(* IEC 61131-3 sources: SortJet_MasterSPS_Aufbau.fbsproj/07_Auftragsverwaltung/Job_Stationen.prg.st^, 8 files *)

(* ---- Auftraege.act.st ---- *)
(* METADATA
{
	"v3Meta": {
		"objectGuid": "798febcb-6f60-456b-b36c-821ba17e31fa"
	}
}
*)
ACTION Auftraege
//-------------------------------------------------------------------------------------------------
// AUFTRAEGE: M_SB0_MMI_SortierungInputInQueue
//-------------------------------------------------------------------------------------------------
(* Hinweis:
   - Anlegetische \ Anlegewaende \ etc. mit einem Auftrag versehen
*)
IF ( M_SB0_MMI_SortierungInputInQueue ) THEN

  CASE tMmi2SpsInfo.wSortierungsInputInQueueStationNr OF

    cERSTE_STATION..cLETZTE_STATION:
      AuftragsSpeicherWand[tMmi2SpsInfo.wSortierungsInputInQueueStationNr, cWAND_1].NeuerAuftrag.rAuftragsHoehe       := tMmi2SpsInfo.rInputInQueueHoehe;
      AuftragsSpeicherWand[tMmi2SpsInfo.wSortierungsInputInQueueStationNr, cWAND_1].NeuerAuftrag.rAuftragsLaenge      := tMmi2SpsInfo.rInputInQueueLaenge;
      AuftragsSpeicherWand[tMmi2SpsInfo.wSortierungsInputInQueueStationNr, cWAND_1].NeuerAuftrag.rAuftragsDicke       := tMmi2SpsInfo.rInputInQueueDicke;
      AuftragsSpeicherWand[tMmi2SpsInfo.wSortierungsInputInQueueStationNr, cWAND_1].NeuerAuftrag.bLetzteScheibe       := 1;
      AuftragsSpeicherWand[tMmi2SpsInfo.wSortierungsInputInQueueStationNr, cWAND_1].NeuerAuftrag.wStationsNr          := tMmi2SpsInfo.wSortierungsInputInQueueStationNr;
      AuftragsSpeicherWand[tMmi2SpsInfo.wSortierungsInputInQueueStationNr, cWAND_1].NeuerAuftrag.wTransferwand        := tMmi2SpsInfo.wSlotZielStation;
      AuftragsSpeicherWand[tMmi2SpsInfo.wSortierungsInputInQueueStationNr, cWAND_1].NeuerAuftrag.wAnzahlScheiben      := 1; // es ist immer nur eine Scheibe anzulegen !
      AuftragsSpeicherWand[tMmi2SpsInfo.wSortierungsInputInQueueStationNr, cWAND_1].NeuerAuftrag.bErsteScheibe        := 1;
      AuftragsSpeicherWand[tMmi2SpsInfo.wSortierungsInputInQueueStationNr, cWAND_1].NeuerAuftrag.bModell              := tMmi2SpsInfo.wModellStatus.0;
      AuftragsSpeicherWand[tMmi2SpsInfo.wSortierungsInputInQueueStationNr, cWAND_1].NeuerAuftrag.rModellVersatzVorne  := tMmi2SpsInfo.rModellVersatzVorne;
      AuftragsSpeicherWand[tMmi2SpsInfo.wSortierungsInputInQueueStationNr, cWAND_1].NeuerAuftrag.rModellVersatzHinten := tMmi2SpsInfo.rModellversatzHinten;
      AuftragsSpeicherWand[tMmi2SpsInfo.wSortierungsInputInQueueStationNr, cWAND_1].NeuerAuftrag.wTransferstationsNr1 := tMmi2SpsInfo.wSourceTable;

      AuftragsSpeicherWand[tMmi2SpsInfo.wSortierungsInputInQueueStationNr, cWAND_1].NeuerAuftrag.wAuftrag := eStation_Anlegen;
      AuftragsSpeicherWand[tMmi2SpsInfo.wSortierungsInputInQueueStationNr, cWAND_1](bpNeuerAuftrag:=TRUE);

      M_SB0_MMI_SortierungInputInQueue := FALSE;

  END_CASE

END_IF

//-------------------------------------------------------------------------------------------------
// AUFTRAEGE: M_SB0_MMI_SORTIERUNGCANCELQUEUEDATA
//-------------------------------------------------------------------------------------------------
(* Hinweis:
   - Aktiven Auftrag eines Anlegetisches loeschen
*)
IF ( M_SB0_MMI_SORTIERUNGCANCELQUEUEDATA ) THEN

  (* Hinweis:
     - Dieser Auftrag darf nur im Automatik- Betrieb validiert \ bearbeitet werden
       => Sendet die HMI diesen Befehl z.B. im Handbetrieb würde der Merker fuer den Abbruch des Anlegeauftrags gesetzt und beim wechsel in den Automatikbetrieb
          würde der nächste Auftrag dann geloescht bzw. abgebrochen und damit verworfen.
       WICHTIG:
     - Sicherstellen das die Stationen diesem Automatikkreis auch angehoehren
  *)
  CASE tMmi2SpsInfo.wDeleteStationNr OF

    cERSTE_STATION..cLETZTE_STATION:
      IF NOT AutomatikAktiv(tMmi2SpsInfo.wDeleteStationNr) THEN
        M_SB0_MMI_SORTIERUNGCANCELQUEUEDATA := FALSE;
      ELSE

        IF ( AuftragsdatenWand[tMmi2SpsInfo.wDeleteStationNr, cWAND_1].wAuftrag = eStation_Anlegen ) THEN
          AuftragsdatenWand[tMmi2SpsInfo.wDeleteStationNr, cWAND_1].wAuftrag := eStation_Kein_Auftrag;
          Anlegen[tMmi2SpsInfo.wDeleteStationNr, cWAND_1](bpReset:=TRUE);
        ELSIF ( AuftragsdatenWand[tMmi2SpsInfo.wDeleteStationNr, cWAND_1].wAuftrag = eStation_Hoehenmessung ) THEN
          AuftragsdatenWand[tMmi2SpsInfo.wDeleteStationNr, cWAND_1].wAuftrag := eStation_Kein_Auftrag;
          Glashoehenmessung[tMmi2SpsInfo.wDeleteStationNr, cWAND_1](bpReset:=TRUE);
        ELSIF ( AuftragsdatenWand[tMmi2SpsInfo.wDeleteStationNr, cWAND_1].wAuftrag = eStation_Messfahrt ) THEN
          AuftragsdatenWand[tMmi2SpsInfo.wDeleteStationNr, cWAND_1].wAuftrag := eStation_Kein_Auftrag;
          Glaslaengenmessung[tMmi2SpsInfo.wDeleteStationNr, cWAND_1](bpReset:=TRUE);
        ELSE
          abpAbbruchAnlegeauftrag[tMmi2SpsInfo.wDeleteStationNr] := TRUE;
        END_IF

        M_SB0_MMI_SORTIERUNGCANCELQUEUEDATA := FALSE;

      END_IF

  END_CASE

END_IF

//-------------------------------------------------------------------------------------------------
// AUFTRAG: M_SB0_MMI_SHEET_ORDER_STATION
//-------------------------------------------------------------------------------------------------
(* Hinweis:
   - -
*)
IF ( M_SB0_MMI_SHEET_ORDER_STATION ) THEN

  IF ( tMmi2SpsInfo.wAuftragsWand = 0 ) THEN // WORKAROUND MMI
    tMmi2SpsInfo.wAuftragsWand := 1;
  END_IF
  IF ( tMmi2SpsInfo.wTransferwand = 0 ) THEN // WORKAROUND MMI
    tMmi2SpsInfo.wTransferwand := 1;
  END_IF

  CASE tMmi2SpsInfo.wStationsNr OF

    cERSTE_STATION..cLETZTE_STATION:
      AuftragsSpeicherWand[tMmi2SpsInfo.wStationsNr, tMmi2SpsInfo.wAuftragsWand].NeuerAuftrag.bModell                 := FALSE;

      AuftragsSpeicherWand[tMmi2SpsInfo.wStationsNr, tMmi2SpsInfo.wAuftragsWand].NeuerAuftrag.wStationsNr             := tMmi2SpsInfo.wStationsNr;          // Stationswand der Quellstation
      AuftragsSpeicherWand[tMmi2SpsInfo.wStationsNr, tMmi2SpsInfo.wAuftragsWand].NeuerAuftrag.wStationsWand           := tMmi2SpsInfo.wAuftragsWand;        // Stationswand der Quellstation
      AuftragsSpeicherWand[tMmi2SpsInfo.wStationsNr, tMmi2SpsInfo.wAuftragsWand].NeuerAuftrag.rStationsZielposition   := tMmi2SpsInfo.rStationsPosition;    // Stationsposition der Quellstation
      AuftragsSpeicherWand[tMmi2SpsInfo.wStationsNr, tMmi2SpsInfo.wAuftragsWand].NeuerAuftrag.rAuftragsLaenge         := tMmi2SpsInfo.rAuftragsLaenge;      // Länge der Scheibe/Batch
      AuftragsSpeicherWand[tMmi2SpsInfo.wStationsNr, tMmi2SpsInfo.wAuftragsWand].NeuerAuftrag.rAuftragsHoehe          := tMmi2SpsInfo.rAuftragsHoehe;       // Höhe der Scheibe/Batch
      AuftragsSpeicherWand[tMmi2SpsInfo.wStationsNr, tMmi2SpsInfo.wAuftragsWand].NeuerAuftrag.rAuftragsDicke          := tMmi2SpsInfo.rAuftragsDicke;       // Dicke der Scheibe/Batch
      AuftragsSpeicherWand[tMmi2SpsInfo.wStationsNr, tMmi2SpsInfo.wAuftragsWand].NeuerAuftrag.wErsteLetzteScheibe     := tMmi2SpsInfo.wErsteLetzteScheibe;  // Kennzeichnung Erste und Letzte Scheibe
      AuftragsSpeicherWand[tMmi2SpsInfo.wStationsNr, tMmi2SpsInfo.wAuftragsWand].NeuerAuftrag.wAnzahlScheiben         := tMmi2SpsInfo.wAnzahlScheiben;      // Anzahl der Scheiben
      AuftragsSpeicherWand[tMmi2SpsInfo.wStationsNr, tMmi2SpsInfo.wAuftragsWand].NeuerAuftrag.wTransferstationsNr1    := tMmi2SpsInfo.wTransferstationsNr1; // Stationsnummer der Zielstation 1
      AuftragsSpeicherWand[tMmi2SpsInfo.wStationsNr, tMmi2SpsInfo.wAuftragsWand].NeuerAuftrag.wTransferstationsNr2    := tMmi2SpsInfo.wTransferstationsNr2; // Stationsnummer der Zielstation 2
      AuftragsSpeicherWand[tMmi2SpsInfo.wStationsNr, tMmi2SpsInfo.wAuftragsWand].NeuerAuftrag.rTransferposition1      := tMmi2SpsInfo.rTransferposition1;   // Stationsposition der Zielstation 1
      AuftragsSpeicherWand[tMmi2SpsInfo.wStationsNr, tMmi2SpsInfo.wAuftragsWand].NeuerAuftrag.rTransferposition2      := tMmi2SpsInfo.rTransferposition2;   // Stationsposition der Zielstation 2
      AuftragsSpeicherWand[tMmi2SpsInfo.wStationsNr, tMmi2SpsInfo.wAuftragsWand].NeuerAuftrag.wTransferwand           := tMmi2SpsInfo.wTransferwand;        // Stationswand der Zielstationen
      AuftragsSpeicherWand[tMmi2SpsInfo.wStationsNr, tMmi2SpsInfo.wAuftragsWand].NeuerAuftrag.stAuftragsInformationen.wAuftragsInformationen  := tMmi2SpsInfo.wAuftragsTyp;         // Informationen zum Auftrag: Bit 1: Ein-Aus-Transport | Bit 2: Station entladen | Bit 3: Ziel FW | Bit 4-7: Wand entladen | etc.

      AuftragsSpeicherWand[tMmi2SpsInfo.wStationsNr, tMmi2SpsInfo.wAuftragsWand].NeuerAuftrag.rModellVersatzVorne     := tMmi2SpsInfo.rModellVersatzVorne;
      AuftragsSpeicherWand[tMmi2SpsInfo.wStationsNr, tMmi2SpsInfo.wAuftragsWand].NeuerAuftrag.rModellVersatzHinten    := tMmi2SpsInfo.rModellversatzHinten;

      IF ((tMmi2SpsInfo.rModellVersatzVorne > 0) OR (tMmi2SpsInfo.rModellVersatzHinten > 0 ) ) THEN
        AuftragsSpeicherWand[tMmi2SpsInfo.wStationsNr, tMmi2SpsInfo.wAuftragsWand].NeuerAuftrag.bModell              := TRUE;
      END_IF

      (* Hinweis:
         - Zuweisung der Bits "erste" und "letzte" Scheibe
      *)

      ErsteUndLetzteScheibeBits( wpErsteUndLetzteScheibe:= tMmi2SpsInfo.wErsteLetzteScheibe ,
                                 wpLetzteScheibe => wlLetzteScheibe,
                                 wpErsteScheibe  => wlErsteScheibe );

      AuftragsSpeicherWand[tMmi2SpsInfo.wStationsNr, tMmi2SpsInfo.wAuftragsWand].NeuerAuftrag.bLetzteScheibe  := wlLetzteScheibe > 0;  // Stationsposition der Zielstation 2
      AuftragsSpeicherWand[tMmi2SpsInfo.wStationsNr, tMmi2SpsInfo.wAuftragsWand].NeuerAuftrag.bErsteScheibe   := wlErsteScheibe  > 0;  // Stationswand der Zielstationen

      IF ( tMmi2SpsInfo.wAuftragsTyp.0 ) THEN
        AuftragsSpeicherWand[tMmi2SpsInfo.wStationsNr, tMmi2SpsInfo.wAuftragsWand].NeuerAuftrag.wAuftrag := eStation_Austransport;
      ELSE
        AuftragsSpeicherWand[tMmi2SpsInfo.wStationsNr, tMmi2SpsInfo.wAuftragsWand].NeuerAuftrag.wAuftrag := eStation_Eintransport;
      END_IF

      AuftragsSpeicherWand[tMmi2SpsInfo.wStationsNr, tMmi2SpsInfo.wAuftragsWand]( bpNeuerAuftrag := TRUE );

      M_SB0_MMI_SHEET_ORDER_STATION := FALSE;

    cERSTE_FREMDANLAGE_AUSLAUF..cLETZTE_FREMDANLAGE_EINLAUF:
      Job_Fremdanlage.AuftragsSpeicherFremdanlage[tMmi2SpsInfo.wStationsNr].NeuerAuftrag.wStationsNr            := tMmi2SpsInfo.wStationsNr;          // Stationswand der Quellstation
      Job_Fremdanlage.AuftragsSpeicherFremdanlage[tMmi2SpsInfo.wStationsNr].NeuerAuftrag.wStationsWand          := tMmi2SpsInfo.wAuftragsWand;        // Stationswand der Quellstation
      Job_Fremdanlage.AuftragsSpeicherFremdanlage[tMmi2SpsInfo.wStationsNr].NeuerAuftrag.rStationsZielposition  := tMmi2SpsInfo.rStationsPosition;    // Stationsposition der Quellstation
      Job_Fremdanlage.AuftragsSpeicherFremdanlage[tMmi2SpsInfo.wStationsNr].NeuerAuftrag.rAuftragsLaenge        := tMmi2SpsInfo.rAuftragsLaenge;      // Länge der Scheibe/Batch
      Job_Fremdanlage.AuftragsSpeicherFremdanlage[tMmi2SpsInfo.wStationsNr].NeuerAuftrag.rAuftragsHoehe         := tMmi2SpsInfo.rAuftragsHoehe;       // Höhe der Scheibe/Batch
      Job_Fremdanlage.AuftragsSpeicherFremdanlage[tMmi2SpsInfo.wStationsNr].NeuerAuftrag.rAuftragsDicke         := tMmi2SpsInfo.rAuftragsDicke;       // Dicke der Scheibe/Batch
      Job_Fremdanlage.AuftragsSpeicherFremdanlage[tMmi2SpsInfo.wStationsNr].NeuerAuftrag.wErsteLetzteScheibe    := tMmi2SpsInfo.wErsteLetzteScheibe;  // Kennzeichnung Erste und Letzte Scheibe
      Job_Fremdanlage.AuftragsSpeicherFremdanlage[tMmi2SpsInfo.wStationsNr].NeuerAuftrag.wAnzahlScheiben        := tMmi2SpsInfo.wAnzahlScheiben;      // Anzahl der Scheiben
      Job_Fremdanlage.AuftragsSpeicherFremdanlage[tMmi2SpsInfo.wStationsNr].NeuerAuftrag.wTransferstationsNr1   := tMmi2SpsInfo.wTransferstationsNr1; // Stationsnummer der Zielstation 1
      Job_Fremdanlage.AuftragsSpeicherFremdanlage[tMmi2SpsInfo.wStationsNr].NeuerAuftrag.wTransferstationsNr2   := tMmi2SpsInfo.wTransferstationsNr2; // Stationsnummer der Zielstation 2
      Job_Fremdanlage.AuftragsSpeicherFremdanlage[tMmi2SpsInfo.wStationsNr].NeuerAuftrag.rTransferposition1     := tMmi2SpsInfo.rTransferposition1;   // Stationsposition der Zielstation 1
      Job_Fremdanlage.AuftragsSpeicherFremdanlage[tMmi2SpsInfo.wStationsNr].NeuerAuftrag.rTransferposition2     := tMmi2SpsInfo.rTransferposition2;   // Stationsposition der Zielstation 2
      Job_Fremdanlage.AuftragsSpeicherFremdanlage[tMmi2SpsInfo.wStationsNr].NeuerAuftrag.wTransferwand          := tMmi2SpsInfo.wTransferwand;        // Stationswand der Zielstationen
      Job_Fremdanlage.AuftragsSpeicherFremdanlage[tMmi2SpsInfo.wStationsNr].NeuerAuftrag.stAuftragsInformationen.wAuftragsInformationen := tMmi2SpsInfo.wAuftragsTyp;         // Informationen zum Auftrag: Bit 1: Ein-Aus-Transport | Bit 2: Station entladen | Bit 3: Ziel FW | Bit 4-7: Wand entladen | etc.

      Job_Fremdanlage.AuftragsSpeicherFremdanlage[tMmi2SpsInfo.wStationsNr].NeuerAuftrag.rModellVersatzVorne  := tMmi2SpsInfo.rModellVersatzVorne;
      Job_Fremdanlage.AuftragsSpeicherFremdanlage[tMmi2SpsInfo.wStationsNr].NeuerAuftrag.rModellVersatzHinten := tMmi2SpsInfo.rModellversatzHinten;

      IF ((tMmi2SpsInfo.rModellVersatzVorne > 0) OR (tMmi2SpsInfo.rModellVersatzHinten > 0 ) ) THEN
        Job_Fremdanlage.AuftragsSpeicherFremdanlage[tMmi2SpsInfo.wStationsNr].NeuerAuftrag.bModell              := TRUE;
      END_IF

      (* Hinweis:
         - Zuweisung der Bits "erste" und "letzte" Scheibe
      *)
      ErsteUndLetzteScheibeBits( wpErsteUndLetzteScheibe:= tMmi2SpsInfo.wErsteLetzteScheibe ,
                                 wpLetzteScheibe => wlLetzteScheibe,
                                 wpErsteScheibe  => wlErsteScheibe );

      Job_Fremdanlage.AuftragsSpeicherFremdanlage[tMmi2SpsInfo.wStationsNr].NeuerAuftrag.bLetzteScheibe  := wlLetzteScheibe > 0;  // Stationsposition der Zielstation 2
      Job_Fremdanlage.AuftragsSpeicherFremdanlage[tMmi2SpsInfo.wStationsNr].NeuerAuftrag.bErsteScheibe   := wlErsteScheibe  > 0;  // Stationswand der Zielstationen

      IF ( tMmi2SpsInfo.wAuftragsTyp.0 ) THEN
        Job_Fremdanlage.AuftragsSpeicherFremdanlage[tMmi2SpsInfo.wStationsNr].NeuerAuftrag.wAuftrag := eStation_Austransport;
      ELSE
        Job_Fremdanlage.AuftragsSpeicherFremdanlage[tMmi2SpsInfo.wStationsNr].NeuerAuftrag.wAuftrag := eStation_Eintransport;
      END_IF

      Job_Fremdanlage.AuftragsSpeicherFremdanlage[tMmi2SpsInfo.wStationsNr]( bpNeuerAuftrag := TRUE );

      M_SB0_MMI_SHEET_ORDER_STATION := FALSE;

    ELSE

      M_SB0_MMI_SHEET_ORDER_STATION := FALSE;

      wpgFehlerdaten[0] := tMmi2SpsInfo.wStationsNr;
      wpgFehlerdaten[1] := tMmi2SpsInfo.wAuftragsWand;
      SpsError( eFehler_Station,
                cMELDUNG_AUFTRAGSDATEN_UNGUELTIGE_STATION,
                tMmi2SpsInfo.wStationsNr,
                AutomatikkreisBestimmen(tMmi2SpsInfo.wStationsNr),
                wpgFehlerdaten );

  END_CASE

END_IF

//-------------------------------------------------------------------------------------------------
// AUFTRAG: M_SB0_MMI_MEASSURERESULT
//-------------------------------------------------------------------------------------------------
(* Hinweis:
   - Scheibeneinlauffreigabe für Anlegetisch
     => Gilt fuer Stationen mit einem Scanner
*)
IF ( M_SB0_MMI_MEASSURERESULT ) THEN

  M_SB0_MMI_MEASSURERESULT := FALSE;

  CASE (tMmi2SpsInfo.wMmiNummerAnlegeStation) OF

    cERSTE_STATION..cLETZTE_STATION:
      ;
    //Anlegewand202.bpFreigabeScheibe      := (tMmi2SpsInfo.wFreigabe = 1);
    //Anlegewand202.bpKeineFreigabeScheibe := (tMmi2SpsInfo.wFreigabe = 0);

    ELSE
      wpgFehlerdaten[0]:= tMmi2SpsInfo.wMmiNummerAnlegeStation;
      wpgFehlerdaten[1]:= tMmi2SpsInfo.wFreigabeStation;
      SpsError( eFehler_Station,
                cMELDUNG_SCANNER_NACHRICHT_FALSCHE_STATION,
                tMmi2SpsInfo.wMmiNummerAnlegeStation,
                AutomatikkreisBestimmen(tMmi2SpsInfo.wMmiNummerAnlegeStation),
                wpgFehlerdaten );

  END_CASE

END_IF

//-------------------------------------------------------------------------------------------------
// AUFTRAG: M_SB0_MMI_STATIONSTATUS
//-------------------------------------------------------------------------------------------------
IF ( M_SB0_MMI_STATIONSTATUS ) THEN

  M_SB0_MMI_STATIONSTATUS := FALSE;

  CASE tMmi2SpsInfo.wStationsNummer OF

    // -------------------------------------------------------------------
    cERSTE_STATION..cLETZTE_STATION:
      (* Hinweis:
         - Aktivieren / Deaktivieren der Station
      *)
      starrStationBasisParameter[tMmi2SpsInfo.wStationsNummer].stMKs.bDeaktivieren := ( NOT tMmi2SpsInfo.wStationsStatusWord7.0 );

    // -------------------------------------------------------------------
    cERSTES_SHUTTLE..cLETZTES_SHUTTLE:
      (* Hinweis:
         - Aktivieren / Deaktivieren der Station
      *)
      starrShuttleBasisParameter[tMmi2SpsInfo.wStationsNummer].stMKs.bDeaktivieren := ( NOT tMmi2SpsInfo.wStationsStatusWord7.0 );

    // -------------------------------------------------------------------
    cERSTES_TRANSFERSHUTTLE..cLETZTES_TRANSFERSHUTTLE:
      (* Hinweis:
         - Aktivieren / Deaktivieren der Station
      *)
      starrTransfershuttleBasisParameter[tMmi2SpsInfo.wStationsNummer].stMKs.bDeaktivieren := ( NOT tMmi2SpsInfo.wStationsStatusWord7.0 );

    // -------------------------------------------------------------------
    cERSTE_FAECHERWAGENSTATIONS_NR..cLETZTE_FAECHERWAGENSTATIONS_NR:
      (* Hinweis:
         - Aktivieren / Deaktivieren der Station
      *)
      starrFaecherwagenBasisParameter[tMmi2SpsInfo.wStationsNummer].stMKs.bDeaktivieren := ( NOT tMmi2SpsInfo.wStationsStatusWord7.0 );
      aFaecherwagenstation[tMmi2SpsInfo.wStationsNummer].wRFID_Nummer_Schreiben := tMmi2SpsInfo.wStationsStatusWord8;

      // Statuswort 1 Bit 0: bei Faecherwagenstationen loest es den Sicherheitskreis-Reset der Station aus
      // (Sicherheitsrelais der Station quittieren)
      IF ( tMmi2SpsInfo.wStationsStatusWord1.0 ) THEN
        aFaecherwagenstation[tMmi2SpsInfo.wStationsNummer].bStarteSicherheitskreisReset := TRUE;
      END_IF

    // -------------------------------------------------------------------
    ELSE
      wpgFehlerdaten[0] := tMmi2SpsInfo.wStationsNummer;
      wpgFehlerdaten[1] := tMmi2SpsInfo.wStationsStatusWord5;
      SpsHinweis( eFehler_Mmi,
                  cMELDUNG_MMI_AUFTRAGSDATEN_UNGUELTIGE_STATIONSNUMMER,
                  0,
                  AutomatikkreisBestimmen(0),
                  wpgFehlerdaten );

  END_CASE

END_IF

//-------------------------------------------------------------------------------------------------
// AUFTRAG: M_SB0_MMI_REQUESTTILTSTATION
//-------------------------------------------------------------------------------------------------

(* Hinweis:
   - Auftrag zum leeren einer Station (Starten eines Austransports)
*)
IF ( M_SB0_MMI_REQUESTTILTSTATION ) THEN

  CASE tMmi2SpsInfo.wSortierungsInputSwingStationNr OF

    cERSTE_STATION..cLETZTE_STATION:
      AuftragsSpeicherWand[tMmi2SpsInfo.wSortierungsInputSwingStationNr, cWAND_1].NeuerAuftrag.wAuftrag      := eStation_Vortransport;
      AuftragsSpeicherWand[tMmi2SpsInfo.wSortierungsInputSwingStationNr, cWAND_1].NeuerAuftrag.wStationsNr   := tMmi2SpsInfo.wSortierungsInputSwingStationNr;
      AuftragsSpeicherWand[tMmi2SpsInfo.wSortierungsInputSwingStationNr, cWAND_1].NeuerAuftrag.wStationsWand := cWAND_1;
      AuftragsSpeicherWand[tMmi2SpsInfo.wSortierungsInputSwingStationNr, cWAND_1]( bpNeuerAuftrag := TRUE );

    ELSE
      wpgFehlerdaten[0] := tMmi2SpsInfo.wSortierungsInputSwingStationNr;
      SpsHinweis( eFehler_Mmi,
                  cMELDUNG_MMI_AUFTRAGSDATEN_UNGUELTIGE_STATIONSNUMMER,
                  0,
                  AutomatikkreisBestimmen(0),
                  wpgFehlerdaten );

  END_CASE

  M_SB0_MMI_REQUESTTILTSTATION := FALSE;

END_IF
END_ACTION

(* ---- Auftragsverwaltung.act.st ---- *)
(* METADATA
{
	"v3Meta": {
		"objectGuid": "ab37f234-5c30-423e-82fd-562034963c76"
	}
}
*)
ACTION Auftragsverwaltung
//-------------------------------------------------------------------------------------------------
// BAUSTEIN: AUFTRAGSVERWALTUNG
//-------------------------------------------------------------------------------------------------
FOR wlIndex := cERSTE_STATION TO cLETZTE_STATION DO

  AuftragsSpeicherStation[wlIndex]();

  IF AuftragsSpeicherStation[wlIndex].bpAuftragverfuegbar
     AND ( AuftragsdatenStation[wlIndex].wAuftrag = eStation_Kein_Auftrag
           OR AuftragsdatenStation[wlIndex].wAuftrag = eStation_Belegt
           OR AuftragsdatenStation[wlIndex].wAuftrag = eStation_Warte_Auf_Eintransport )
  THEN
    AuftragsSpeicherStation[wlIndex].bpNaechsterAuftrag := TRUE;
    AuftragsSpeicherStation[wlIndex]();
    AuftragsdatenStation[wlIndex] := AuftragsSpeicherStation[wlIndex].AktAuftrag;
  END_IF

  FOR wlIndexWand := cWAND_1 TO cANZAHL_WAENDE DO

    AuftragsSpeicherWand[wlIndex, wlIndexWand]();

    IF AuftragsSpeicherWand[wlIndex, wlIndexWand].bpAuftragverfuegbar
       AND ( AuftragsdatenWand[wlIndex, wlIndexWand].wAuftrag = eStation_Kein_Auftrag
             OR AuftragsdatenWand[wlIndex, wlIndexWand].wAuftrag = eStation_Belegt
             OR AuftragsdatenWand[wlIndex, wlIndexWand].wAuftrag = eStation_Warte_Auf_Eintransport
             OR AuftragsdatenWand[wlIndex, wlIndexWand].wAuftrag = eStation_Warte_Auf_Austransport  )
    THEN
      AuftragsSpeicherWand[wlIndex, wlIndexWand].bpNaechsterAuftrag := TRUE;
      AuftragsSpeicherWand[wlIndex, wlIndexWand]();
      AuftragsdatenWand[wlIndex, wlIndexWand] := AuftragsSpeicherWand[wlIndex, wlIndexWand].AktAuftrag;
    END_IF

  END_FOR

END_FOR
END_ACTION

(* ---- Reset.act.st ---- *)
(* METADATA
{
	"v3Meta": {
		"objectGuid": "37f6c3a9-3bba-4d57-9c53-2ef1e7be2c3a"
	}
}
*)
ACTION Reset
//-------------------------------------------------------------------------------------------------
// AKTION: RESET
//-------------------------------------------------------------------------------------------------

FOR wlIndexReset := cERSTER_AUTOMATIKKREIS TO cLETZTER_AUTOMATIKKREIS DO

  IF ( abpReset[wlIndexReset] ) THEN

    abpReset[wlIndexReset] := FALSE;
    abpFehler[wlIndexReset] := FALSE;

    FOR wlIndex := cERSTE_STATION TO cLETZTE_STATION DO

      IF StationInAutomatikkreis(starrStationBasisParameter[wlIndex].stMKs.eaAutomatikkreis, wlIndexReset) THEN

        abpAbbruchAnlegeauftrag[wlIndex] := FALSE;

        AuftragsSpeicherStation[wlIndex].bpReset := TRUE;
        AuftragsSpeicherStation[wlIndex]();

        AuftragsdatenStation[wlIndex].wAuftrag := eStation_Kein_Auftrag;

        starrStationBasisParameter[wlIndex].bReset := TRUE;

        FOR wlIndexWand := cWAND_1 TO cANZAHL_WAENDE DO

          AuftragsSpeicherWand[wlIndex,wlIndexWand].bpReset := TRUE;
          AuftragsSpeicherWand[wlIndex,wlIndexWand]();

          AuftragsdatenWand[wlIndex, wlIndexWand].wAuftrag := eStation_Kein_Auftrag;

          ailScheibenZuQuittierenEintransport[wlIndex, wlIndexWand] := 0;
          ailScheibenZuQuittierenAustransport[wlIndex, wlIndexWand] := 0;

          ablMerkerLetzteScheibeStation[wlIndex, wlIndexWand] := FALSE;

          ablFreigabeZurParalleleBausteinAnsteuerung[wlIndex,wlIndexWand] := FALSE;
          abpStarteParalleleBausteinAnsteuerung[wlIndex, wlIndexWand]     := FALSE;

        END_FOR

      END_IF

    END_FOR

  END_IF

END_FOR
END_ACTION

(* ---- Schnittstelle_Stationen.act.st ---- *)
(* METADATA
{
	"v3Meta": {
		"objectGuid": "2f0e1e2b-c489-43f6-919f-1d41b03fa1f2"
	}
}
*)
ACTION Schnittstelle_Stationen
//-------------------------------------------------------------------------------------------------
// SCHNITTSTELLE ZWISCHEN DEN STATIONEN
//-------------------------------------------------------------------------------------------------

//  KOPPLUNGEN

//starrFremdanlageEinlaufStationBasisParameter[501].InGlasTransportNachfolger[cWAND_1] := starrStationBasisParameter[cSTATION_201].OutGlasTransport[cWAND_1];
//starrStationBasisParameter[cSTATION_201].InGlasTransportVorgaenger[cWAND_1] := starrFremdanlageEinlaufStationBasisParameter[501].OutGlasTransport[cWAND_1];

FOR wlIndex := cERSTE_STATION TO cLETZTE_FREMDANLAGE_EINLAUF DO

  // Struktur für die Zielstation der Kopplung finden
  stLokaleKopplungZielStation REF= getBasis(wlIndex);

  IF __ISVALIDREF(stLokaleKopplungZielStation) THEN

    // Kopplung Vorgänger
    stLokaleKopplungsStation REF= getBasis(stLokaleKopplungZielStation.stMKs.stSchnittstellendaten.wVorgaengerStation);

    IF __ISVALIDREF(stLokaleKopplungsStation) THEN
      FOR wlIndexWand := cWAND_1 TO cANZAHL_WAENDE DO
        stLokaleKopplungZielStation.InGlasTransportVorgaenger[wlIndexWand] := stLokaleKopplungsStation.OutGlasTransport[cWAND_1];
      END_FOR
    END_IF

    // Kopplung Nachfolger
    stLokaleKopplungsStation REF= getBasis(stLokaleKopplungZielStation.stMKs.stSchnittstellendaten.wNachfolgerStation);

    IF __ISVALIDREF(stLokaleKopplungsStation) THEN
      FOR wlIndexWand := cWAND_1 TO cANZAHL_WAENDE DO
        stLokaleKopplungZielStation.InGlasTransportNachfolger[wlIndexWand] := stLokaleKopplungsStation.OutGlasTransport[cWAND_1];
      END_FOR
    END_IF

  END_IF

END_FOR
END_ACTION

(* ---- Station.meth.st ---- *)
(* METADATA
{
	"v3Meta": {
		"objectGuid": "6e43b8d4-0bae-4a3f-b309-8e06ab9993e4"
	}
}
*)
METHOD INTERNAL Station
VAR_INPUT
  wStation : WORD;
  wWand    : WORD;
END_VAR

// ****************************************************9*********************************************
// STEUERUNG: ANLEGEN
// *************************************************************************************************

IF ( AuftragsdatenWand[wStation, wWand].wAuftrag = eStation_Anlegen ) THEN
  (* Hinweis:
     - Aufruf der Schrittkette
  *)
  Anlegen[wStation, wWand]( Auftragsdaten := AuftragsdatenWand[wStation, wWand], bpAbbruchAnlegeauftrag := abpAbbruchAnlegeauftrag[wStation], wStation := wStation);
  (* Hinweis:
     - Abschluss der Schrittkette
  *)
  IF Anlegen[wStation, wWand].bpDone THEN
    abpAbbruchAnlegeauftrag[wStation] := FALSE;
    AuftragsdatenWand[wStation, wWand] := Anlegen[wStation, wWand].Auftragsdaten;
    Anlegen[wStation, wWand](bpReset := TRUE);
  END_IF
  (* Hinweis:
     - Fehler-Auswertung
  *)
  ablFehler[wStation, wWand] := Anlegen[wStation, wWand].bpFehler;
  IF rtlFehler[wStation, wWand].Q THEN
    AutomatikFehlerSetzen(starrStationBasisParameter[wStation].stMKs.eaAutomatikkreis, abpFehler);
  END_IF
ELSE
  (* Hinweis:
     - Reset der Schrittkette
  *)
  IF ( Anlegen[wStation, wWand].steplSchritt > STEP_0_E ) THEN
    Anlegen[wStation, wWand](bpReset := TRUE);
  END_IF
END_IF

// ****************************************************9*********************************************
// STEUERUNG: ABNEHMEN
// *************************************************************************************************

IF ( AuftragsdatenWand[wStation, wWand].wAuftrag = eStation_Abnehmen ) THEN
  (* Hinweis:
     - Aufruf der Schrittkette
  *)
  Abnehmen[wStation, wWand]( Auftragsdaten := AuftragsdatenWand[wStation, wWand], wStation := wStation);
  (* Hinweis:
     - Abschluss der Schrittkette
  *)
  IF Abnehmen[wStation, wWand].bpDone THEN
    abpAbbruchAnlegeauftrag[wStation] := FALSE;
    AuftragsdatenWand[wStation, wWand] := Abnehmen[wStation, wWand].Auftragsdaten;
    Abnehmen[wStation, wWand](bpReset := TRUE);
  END_IF
  (* Hinweis:
     - Fehler-Auswertung
  *)
  ablFehler[wStation, wWand] := Abnehmen[wStation, wWand].bpFehler;
  IF rtlFehler[wStation, wWand].Q THEN
    AutomatikFehlerSetzen(starrStationBasisParameter[wStation].stMKs.eaAutomatikkreis, abpFehler);
  END_IF
ELSE
  (* Hinweis:
     - Reset der Schrittkette
  *)
  IF ( Abnehmen[wStation, wWand].steplSchritt > STEP_0_E ) THEN
    Abnehmen[wStation, wWand](bpReset := TRUE);
  END_IF
END_IF

// ****************************************************9*********************************************
// STEUERUNG: HÖHENMESSUNG
// *************************************************************************************************

IF ( AuftragsdatenWand[wStation, wWand].wAuftrag = eStation_Hoehenmessung ) THEN
  (* Hinweis:
     - Aufruf der Schrittkette
  *)
  Glashoehenmessung[wStation, wWand]( Auftragsdaten := AuftragsdatenWand[wStation, wWand], wStation := wStation, bpAbbruchAnlegeauftrag := abpAbbruchAnlegeauftrag[wStation]);
  (* Hinweis:
     - Abschluss der Schrittkette
  *)
  IF Glashoehenmessung[wStation, wWand].bpDone THEN
    abpAbbruchAnlegeauftrag[wStation] := FALSE;
    AuftragsdatenWand[wStation, wWand] := Glashoehenmessung[wStation, wWand].Auftragsdaten;
    Glashoehenmessung[wStation, wWand](bpReset := TRUE);
  END_IF
  (* Hinweis:
     - Fehler-Auswertung
  *)
  ablFehler[wStation, wWand] := Glashoehenmessung[wStation, wWand].bpFehler;
  IF rtlFehler[wStation, wWand].Q THEN
    AutomatikFehlerSetzen(starrStationBasisParameter[wStation].stMKs.eaAutomatikkreis, abpFehler);
  END_IF
ELSE
  (* Hinweis:
     - Reset der Schrittkette
  *)
  IF ( Glashoehenmessung[wStation, wWand].steplSchritt > STEP_0_E ) THEN
    Glashoehenmessung[wStation, wWand](bpReset := TRUE);
  END_IF
END_IF

// ****************************************************9*********************************************
// STEUERUNG: LÄNGENMESSUNG
// *************************************************************************************************

IF ( AuftragsdatenWand[wStation, wWand].wAuftrag = eStation_Messfahrt ) THEN
  (* Hinweis:
     - Aufruf der Schrittkette
  *)
  Glaslaengenmessung[wStation, wWand]( Auftragsdaten := AuftragsdatenWand[wStation, wWand], wStation := wStation, bpAbbruchAnlegeauftrag := abpAbbruchAnlegeauftrag[wStation] );
  (* Hinweis:
     - Abschluss der Schrittkette
  *)
  IF Glaslaengenmessung[wStation, wWand].bpDone THEN
    abpAbbruchAnlegeauftrag[wStation] := FALSE;
    AuftragsdatenWand[wStation, wWand] := Glaslaengenmessung[wStation, wWand].Auftragsdaten;
    Glaslaengenmessung[wStation, wWand](bpReset := TRUE);
  END_IF
  (* Hinweis:
     - Fehler-Auswertung
  *)
  ablFehler[wStation, wWand] := Glaslaengenmessung[wStation, wWand].bpFehler;
  IF rtlFehler[wStation, wWand].Q THEN
    AutomatikFehlerSetzen(starrStationBasisParameter[wStation].stMKs.eaAutomatikkreis, abpFehler);
  END_IF
ELSE
  (* Hinweis:
     - Reset der Schrittkette
  *)
  IF ( Glaslaengenmessung[wStation, wWand].steplSchritt > STEP_0_E ) THEN
    Glaslaengenmessung[wStation, wWand](bpReset := TRUE);
  END_IF
END_IF

// ****************************************************9*********************************************
// STEUERUNG: Eintransport
// *************************************************************************************************

IF ( AuftragsdatenWand[wStation, wWand].wAuftrag = eStation_Eintransport ) THEN
  (* Hinweis:
     - Aufruf der Schrittkette
  *)
  Eintransport[wStation, wWand]( Auftragsdaten := AuftragsdatenWand[wStation, wWand], wStation := wStation, wWand := wWand);
  (* Hinweis:
     - Abschluss der Schrittkette
  *)
  IF Eintransport[wStation, wWand].bpDone THEN
    AuftragsdatenWand[wStation, wWand] := Eintransport[wStation, wWand].Auftragsdaten;
    Eintransport[wStation, wWand](bpReset := TRUE);
  END_IF
  (* Hinweis:
     - Fehler-Auswertung
  *)
  ablFehler[wStation, wWand] := Eintransport[wStation, wWand].bpFehler;
  IF rtlFehler[wStation, wWand].Q THEN
    AutomatikFehlerSetzen(starrStationBasisParameter[wStation].stMKs.eaAutomatikkreis, abpFehler);
  END_IF
ELSE
  (* Hinweis:
     - Reset der Schrittkette
  *)
  IF ( Eintransport[wStation, wWand].steplSchritt > STEP_0_E ) THEN
    Eintransport[wStation, wWand](bpReset := TRUE);
  END_IF
END_IF

// ****************************************************9*********************************************
// STEUERUNG: AUSTRANSPORT
// *************************************************************************************************

IF ( AuftragsdatenWand[wStation, wWand].wAuftrag = eStation_Austransport ) THEN
  (* Hinweis:
     - Aufruf der Schrittkette
  *)
  Austransport[wStation, wWand]( Auftragsdaten := AuftragsdatenWand[wStation, wWand], wStation := wStation, wWand := wWand);
  (* Hinweis:
     - Abschluss der Schrittkette
  *)
  IF Austransport[wStation, wWand].bpDone THEN
    AuftragsdatenWand[wStation, wWand] := Austransport[wStation, wWand].Auftragsdaten;
    Austransport[wStation, wWand](bpReset := TRUE);
  END_IF
  (* Hinweis:
     - Fehler-Auswertung
  *)
  ablFehler[wStation, wWand] := Austransport[wStation, wWand].bpFehler;
  IF rtlFehler[wStation, wWand].Q THEN
    AutomatikFehlerSetzen(starrStationBasisParameter[wStation].stMKs.eaAutomatikkreis, abpFehler);
  END_IF
ELSE
  (* Hinweis:
     - Reset der Schrittkette
  *)
  IF ( Austransport[wStation, wWand].steplSchritt > STEP_0_E ) THEN
    Austransport[wStation, wWand](bpReset := TRUE);
  END_IF
END_IF

// ****************************************************9*********************************************
// STEUERUNG: DURCHTRANSPORT
// *************************************************************************************************

IF ( AuftragsdatenWand[wStation, wWand].wAuftrag = eStation_Durchtransport ) THEN
  (* Hinweis:
     - Aufruf der Schrittkette
  *)
  Durchtransport[wStation, wWand]( Auftragsdaten := AuftragsdatenWand[wStation, wWand], wStation := wStation, wWand := wWand);
  (* Hinweis:
     - Abschluss der Schrittkette
  *)
  IF Durchtransport[wStation, wWand].bpDone THEN
    AuftragsdatenWand[wStation, wWand] := Durchtransport[wStation, wWand].Auftragsdaten;
    Durchtransport[wStation, wWand](bpReset := TRUE);
  END_IF
  (* Hinweis:
     - Fehler-Auswertung
  *)
  ablFehler[wStation, wWand] := Durchtransport[wStation, wWand].bpFehler;
  IF rtlFehler[wStation, wWand].Q THEN
    AutomatikFehlerSetzen(starrStationBasisParameter[wStation].stMKs.eaAutomatikkreis, abpFehler);
  END_IF
ELSE
  (* Hinweis:
     - Reset der Schrittkette
  *)
  IF ( Durchtransport[wStation, wWand].steplSchritt > STEP_0_E ) THEN
    Durchtransport[wStation, wWand](bpReset := TRUE);
  END_IF
END_IF

// ****************************************************9*********************************************
// STEUERUNG: Vortransport
// *************************************************************************************************

IF ( AuftragsdatenWand[wStation, wWand].wAuftrag = eStation_Vortransport ) THEN
  (* Hinweis:
     - Aufruf der Schrittkette
  *)
  Vortransport[wStation, wWand]( Auftragsdaten := AuftragsdatenWand[wStation, wWand], wStation := wStation, wWand := wWand);
  (* Hinweis:
     - Abschluss der Schrittkette
  *)
  IF Vortransport[wStation, wWand].bpDone THEN
    AuftragsdatenWand[wStation, wWand] := Vortransport[wStation, wWand].Auftragsdaten;
    Vortransport[wStation, wWand](bpReset := TRUE);
  END_IF
  (* Hinweis:
     - Fehler-Auswertung
  *)
  ablFehler[wStation, wWand] := Vortransport[wStation, wWand].bpFehler;
  IF rtlFehler[wStation, wWand].Q THEN
    AutomatikFehlerSetzen(starrStationBasisParameter[wStation].stMKs.eaAutomatikkreis, abpFehler);
  END_IF
ELSE
  (* Hinweis:
     - Reset der Schrittkette
  *)
  IF ( Vortransport[wStation, wWand].steplSchritt > STEP_0_E ) THEN
    Vortransport[wStation, wWand](bpReset := TRUE);
  END_IF
END_IF

// ****************************************************9*********************************************
// STEUERUNG: TRANSPORTKOPPLUNG
// *************************************************************************************************

IF ( AuftragsdatenWand[wStation, wWand].wAuftrag = eStation_Transportkopplung ) THEN
  (* Hinweis:
     - Aufruf der Schrittkette
  *)
  Transportkopplung[wStation, wWand]( Auftragsdaten := AuftragsdatenWand[wStation, wWand], wStation := wStation, wWand := wWand);
  (* Hinweis:
     - Abschluss der Schrittkette
  *)
  IF Transportkopplung[wStation, wWand].bpDone THEN
    AuftragsdatenWand[wStation, wWand] := Transportkopplung[wStation, wWand].Auftragsdaten;
    Transportkopplung[wStation, wWand](bpReset := TRUE);
  END_IF
  (* Hinweis:
     - Fehler-Auswertung
  *)
  ablFehler[wStation, wWand] := Transportkopplung[wStation, wWand].bpFehler;
  IF rtlFehler[wStation, wWand].Q THEN
    AutomatikFehlerSetzen(starrStationBasisParameter[wStation].stMKs.eaAutomatikkreis, abpFehler);
  END_IF
ELSE
  (* Hinweis:
     - Reset der Schrittkette
  *)
  IF ( Transportkopplung[wStation, wWand].steplSchritt > STEP_0_E ) THEN
    Transportkopplung[wStation, wWand](bpReset := TRUE);
  END_IF
END_IF
// ****************************************************9*********************************************
// STEUERUNG: MESSKOPPLUNG
// *************************************************************************************************

IF ( AuftragsdatenWand[wStation, wWand].wAuftrag = eStation_Messkopplung )
THEN
  (* Hinweis:
     - Aufruf der Schrittkette
  *)
  Messkopplung[wStation, wWand]( Auftragsdaten := AuftragsdatenWand[wStation, wWand], wStation := wStation, wWand := wWand);
  (* Hinweis:
     - Abschluss der Schrittkette
  *)
  IF Transportkopplung[wStation, wWand].bpDone THEN
    AuftragsdatenWand[wStation, wWand] := Messkopplung[wStation, wWand].Auftragsdaten;
    Messkopplung[wStation, wWand](bpReset := TRUE);
  END_IF
  (* Hinweis:
     - Fehler-Auswertung
  *)
  ablFehler[wStation, wWand] := Messkopplung[wStation, wWand].bpFehler;
  IF rtlFehler[wStation, wWand].Q THEN
    AutomatikFehlerSetzen(starrStationBasisParameter[wStation].stMKs.eaAutomatikkreis, abpFehler);
  END_IF
ELSE
  (* Hinweis:
     - Reset der Schrittkette
  *)
  IF ( Messkopplung[wStation, wWand].steplSchritt > STEP_0_E ) THEN
    Messkopplung[wStation, wWand](bpReset := TRUE);
  END_IF
END_IF

// ****************************************************9*********************************************
// STEUERUNG: QUERFAHRT
// *************************************************************************************************

IF ( AuftragsdatenStation[wStation].wAuftrag = eStation_Vorabpositionierung ) THEN
  (* Hinweis:
     - Aufruf der Schrittkette
  *)
  Querfahrt[wStation]( Auftragsdaten := AuftragsdatenStation[wStation], wStation := wStation );
  (* Hinweis:
     - Abschluss der Schrittkette
  *)
  IF Querfahrt[wStation].bpDone THEN
    AuftragsdatenStation[wStation] := Querfahrt[wStation].Auftragsdaten;
    Querfahrt[wStation](bpReset := TRUE);
  END_IF
  (* Hinweis:
     - Fehler-Auswertung
  *)
  ablFehler[wStation, cWAND_1] := Querfahrt[wStation].bpFehler;
  IF rtlFehler[wStation, cWAND_1].Q THEN
    AutomatikFehlerSetzen(starrStationBasisParameter[wStation].stMKs.eaAutomatikkreis, abpFehler);
  END_IF
ELSE
  (* Hinweis:
     - Reset der Schrittkette
  *)
  IF ( Querfahrt[wStation].steplSchritt <> STEP_0_E ) THEN
    Querfahrt[wStation](bpReset := TRUE);
  END_IF
END_IF
END_METHOD

(* ---- Status_Automatikkreis_Start.act.st ---- *)
(* METADATA
{
	"v3Meta": {
		"objectGuid": "48c1475d-7d1e-4064-b68a-f94b7224aadc"
	}
}
*)
ACTION Status_Automatikkreis_Start
//-------------------------------------------------------------------------------------------------
// AKTION: AUFTRAGSSTATUS SETZEN BEIM STARTEN DAS AUTOMATIKMODUS
//-------------------------------------------------------------------------------------------------

FOR wlIndexAutoStart := cERSTER_AUTOMATIKKREIS TO cLETZTER_AUTOMATIKKREIS DO

  rtlStartAutomatik[wlIndexAutoStart](CLK := M_Automatik_Aktiv[wlIndexAutoStart] OR Visu_Start_Auto);

  IF ( rtlStartAutomatik[wlIndexAutoStart].Q ) THEN

    FOR wlIndex := cERSTE_STATION TO cLETZTE_STATION DO
      IF ( StationInAutomatikkreis(starrStationBasisParameter[wlIndex].stMKs.eaAutomatikkreis, wlIndexAutoStart) ) THEN

        FOR wlIndexWand := cWAND_1 TO cANZAHL_WAENDE DO
          Job_Stationen.AuftragsdatenWand[wlIndex, wlIndexWand].wAuftrag := starrStationBasisParameter[wlIndex].pAuftragNachSystemcheck[wlIndexWand];
        END_FOR

      END_IF

    END_FOR

  END_IF

END_FOR
END_ACTION

(* ---- Verfahrfreigabe.act.st ---- *)
(* METADATA
{
	"v3Meta": {
		"objectGuid": "947d4714-9a33-4aa6-8a4d-61239e97d0f5"
	}
}
*)
ACTION Verfahrfreigabe
//-------------------------------------------------------------------------------------------------
// VERFAHRFREIGABE STATIONEN
//-------------------------------------------------------------------------------------------------
(* Hinweis [STATIONEN]:
   - Zurueck des Auftrags  "eStation_Vorabpositionierung" wenn dieser aktiv gewesen ist
     => Verfahrlogik
*)
FOR wlIndex := cERSTE_STATION TO cLETZTE_STATION DO
  IF  ( starrStationBasisParameter[wlIndex].bPositionierAuftragZuruecksetzen ) THEN
    IF ( AuftragsdatenStation[wlIndex].wAuftrag = eStation_Vorabpositionierung ) THEN
      starrStationBasisParameter[wlIndex].bQuittungPositionierungZurueckgesetzt := TRUE;
      AuftragsdatenStation[wlIndex].wAuftrag := eStation_Kein_Auftrag;
    END_IF
  END_IF
END_FOR
END_ACTION

(* ---- Visu.act.st ---- *)
(* METADATA
{
	"v3Meta": {
		"objectGuid": "ba58e9e7-a53f-4b72-9d20-33bd7cca2a1a"
	}
}
*)
ACTION Visu
// *************************************************************************************************
// Daten in das VisoArray kopieren
FOR wlIndex := cERSTE_STATION TO cLETZTE_STATION DO
  VisuAuftragsdaten[wlIndex].eStation := TO_WORD(AuftragsdatenStation[wlIndex].wAuftrag);
  FOR wlIndexWand := cWAND_1 TO cANZAHL_WAENDE DO
    VisuAuftragsdaten[wlIndex].eWand[wlIndexWand] := TO_WORD(AuftragsdatenWand[wlIndex, wlIndexWand].wAuftrag);
  END_FOR
END_FOR
END_ACTION
